(* IEC 61131-3 sources: FibonacciChallenge/Network/FibonacciChallegeNetwork, 1 file *)

(* ---- ONE_FibonacciChallegeNetwork_Table.st ---- *)
#define OBJECTS_CONFIG

FUNCTION GLOBAL TAB ONE_FibonacciChallegeNetwork
-1$UINT, 0$UINT,
0$UINT, 0$UINT,

1$UDINT,
TO_UDINT(3858999192), "FibChallenge", 0$UINT, 0$UINT, 1$UINT,

_NO_ATTR, TO_UDINT(2112812902), "FIBCHALLENGE1",

//Internal connections
0$UDINT,
0$UDINT,
0$UDINT,
0$UDINT,

//Initialization values
0$UDINT,
0$UDINT,

//Symbolic initialization values
0$UDINT,
0$UDINT,

//Initialization of string values
0$UDINT,
0$UDINT,

//Configuration of tasks (RealTime, Cyclic, Background)
0$UDINT,
0$UDINT,

0$UDINT,
1$UDINT,
TO_UDINT(0), (1)$UDINT, 4194303$DINT, 	//FIBCHALLENGE1

0$UDINT,
0$UDINT,

//External connections
0$UDINT,
0$UDINT,

//Magic internal connections
0$UDINT,
0$UDINT,

//Configuration of timeslots of tasks (RealTime, Cyclic)
#ifdef __LSLLDR_TIMESLOTS__
0$UDINT,
0$UDINT,

0$UDINT,
0$UDINT,

#endif //__LSLLDR_TIMESLOTS__

//MultiMaster connections
#ifdef __LSLLDR_MULTIMASTER__
0$UDINT,
0$UDINT,
#endif //__LSLLDR_MULTIMASTER__

//Configuration for task ID (RealTime, CyclicTime)
#ifdef __LSLLDR_TASKID__
"\\\\TASKS2  "
0$UDINT,
0$UDINT,

0$UDINT,
1$UDINT,
(0)$UDINT, 	//FIBCHALLENGE1

0$UDINT,
0$UDINT,

#endif //__LSLLDR_TASKID__

END_FUNCTION
